(* IEC 61131-3 sources: guidance-for-physical-ai-production-designer-on-aws/source/plan2cell/examples/welding_cell_2_small/plc/codesys/robots/robot2/POU, 10 files *)

(* ---- FB_JointAngleEncoder.st ---- *)
(*
 * FB_JointAngleEncoder
 * Device simulator R2 (robot2), cell welding_cell_2_small. Generated by bt2plc 0.1.0.
 *
 * Encodes six KUKA robot joint angles (REAL degrees) into the VASS Option area
 * as scaled fixed-point INTs (0.02 deg per count, big-endian byte order).
 *
 * Encoding per encoding.md:
 *   count = ROUND(angle_deg / 0.02)   clamped to [-32768, +32767]
 *   Byte layout: big-endian (high byte first) in each 2-byte pair
 *
 * Output abyOption = Option area aVassInputData[16..27], 2 bytes per axis
 * (PLC_PRG copies it into the robot -> PLC telegram):
 *   abyOption[0-1]  = bytes 16-17 = A1,  abyOption[2-3]   = bytes 18-19 = A2,
 *   abyOption[4-5]  = bytes 20-21 = A3,  abyOption[6-7]   = bytes 22-23 = A4,
 *   abyOption[8-9]  = bytes 24-25 = A5,  abyOption[10-11] = bytes 26-27 = A6
 *)

FUNCTION_BLOCK FB_JointAngleEncoder
VAR_INPUT
    rA1_deg     : REAL := 0.0;      (* Axis 1 angle in degrees *)
    rA2_deg     : REAL := 0.0;      (* Axis 2 angle in degrees *)
    rA3_deg     : REAL := 0.0;      (* Axis 3 angle in degrees *)
    rA4_deg     : REAL := 0.0;      (* Axis 4 angle in degrees *)
    rA5_deg     : REAL := 0.0;      (* Axis 5 angle in degrees *)
    rA6_deg     : REAL := 0.0;      (* Axis 6 angle in degrees *)
END_VAR

VAR_OUTPUT
    (* Encoded INT values (for monitoring/debug) *)
    iA1_count   : INT;
    iA2_count   : INT;
    iA3_count   : INT;
    iA4_count   : INT;
    iA5_count   : INT;
    iA6_count   : INT;

    (* Option area bytes 16..27 of the robot -> PLC telegram, big-endian A1..A6 *)
    abyOption   : ARRAY[0..11] OF BYTE;
END_VAR

VAR CONSTANT
    SCALE_FACTOR    : REAL := 0.02;     (* degrees per count *)
    INV_SCALE       : REAL := 50.0;     (* 1/0.02 = 50, multiply for speed *)
    COUNT_MAX       : DINT := 32767;
    COUNT_MIN       : DINT := -32768;
END_VAR

VAR
    _arDeg      : ARRAY[1..6] OF REAL;
    _aiCount    : ARRAY[1..6] OF INT;
    _diTemp     : DINT;
    _wTemp      : WORD;
    _i          : INT;
END_VAR

(* ---- FB_PROFIsafe_Simulator.st ---- *)
(*
 * FB_PROFIsafe_Simulator
 * Device simulator R2 (robot2), cell welding_cell_2_small. Generated by bt2plc 0.1.0.
 *
 * Simulates the PROFIsafe protocol layer for the FDIO64 module (Slot 1).
 * In a real KUKA controller, the PROFIsafe stack handles CRC generation,
 * sequence counters, and watchdog monitoring.
 *
 * For simulation purposes, this FB:
 * - Monitors the safe output bytes from the PLC (abySafeOut = copy of GVL_IO.bySafeOut0..7)
 * - Provides a "communication OK" flag
 *
 * IMPORTANT: This does NOT provide real functional safety!
 * It only generates data patterns that allow the PLC's PROFIsafe stack
 * to accept the device as communicating. For real safety testing,
 * you need a certified PROFIsafe device or test equipment.
 *
 * PROFIsafe frame structure per IEC 61784-3-3:
 *   [User Data (8 bytes)] [Status/Control (1 byte)] [CRC (3 bytes)]
 *
 * Status byte bits (F_Input from device):
 *   Bit 0: Toggle bit (alternates each cycle)
 *   Bit 1: Reserved
 *   Bit 2: Data valid
 *   Bit 3-7: Reserved / Sequence counter
 *
 * Control byte bits (F_Output from controller):
 *   Bit 0: Toggle bit
 *   Bit 1: Activate device
 *   Bit 2: Reserved
 *   Bit 3-7: Reserved
 *)

FUNCTION_BLOCK FB_PROFIsafe_Simulator
VAR_INPUT
    bEnable         : BOOL := TRUE;
    dwF_Source_Add  : DWORD := DWORD#1;     (* F_Source_Add from parameterization *)
    dwF_Dest_Add    : DWORD := DWORD#1;     (* F_Dest_Add from parameterization *)
    tF_WD_Time      : TIME := T#500MS;      (* Watchdog time *)
    abySafeOut      : ARRAY[0..7] OF BYTE;  (* Safe outputs PLC -> robot (GVL_IO.bySafeOut0..7) *)
END_VAR

VAR_OUTPUT
    bCommOK         : BOOL;                 (* PROFIsafe communication established *)
    bDataValid      : BOOL;                 (* Safe data is valid *)
    bWatchdogError  : BOOL;                 (* Watchdog timeout *)
END_VAR

VAR
    _bToggleBit     : BOOL;                 (* Toggle bit for sequence *)
    _nSeqCounter    : BYTE;                 (* Sequence counter 0-31 *)
    _nCycleCount    : UDINT;                (* Absolute cycle counter *)

    (* Watchdog *)
    _tonWatchdog    : TON;
    _bPLCSafeActive : BOOL;

    (* CRC calculation helper *)
    _dwCrcSeed      : DWORD;
END_VAR

(* ---- FB_ProgramPlayer.st ---- *)
(*
 * FB_ProgramPlayer
 * Device simulator R2 (robot2), cell welding_cell_2_small, tree bt_1790934549_welding_cell_2_small. Generated by bt2plc 0.1.0.
 *
 * Plays the bt2plc robot program (GVL_Program) for PROD_FOLGE, or a blind joint
 * move to the home pose for HOME_FOLGE. Robot side of the zone protocol, per op k
 * with mask M = GVL_Program.aOps[k].dwZoneMask:
 *   1  wStep := k                          (also for M = 0)
 *   2  if M <> 0: REQUEST := M             (same call / telegram as wStep)
 *   3  if M <> 0: wait (GRANT AND M) = M
 *   4  start delay; trajectory (x rVelScale x override); hold
 *   5  if M <> 0: REQUEST := 0
 *   6  if M <> 0: wait (GRANT AND M) = 0   (4-phase, before the next REQUEST)
 *   7  next op; after the last op: bDone, wStep := 0 (same call)
 *
 * Timing: all times are REAL seconds accumulated from rDt (seconds per call, the
 * device task interval). Motion time advances by rDt * rRate * rVelScale, delay and
 * hold by rDt (the override does not scale dwell times). No TIME() / TON is used.
 * Zero-time transitions fall through within one call (at most N_MAX_TRANSITIONS),
 * but wStep changes at most once per call, so every step is visible to the head PLC.
 * Joints (deg) are linearly interpolated between waypoints and published as rA1..rA6_deg.
 * Abort (bAbort level while busy): REQUEST := 0, wStep := 0, the pose is held.
 * The robot powers up at GVL_Program.arHomeDeg.
 *)

FUNCTION_BLOCK FB_ProgramPlayer
VAR_INPUT
    bStart          : BOOL;                 (* Rising edge: start wJob *)
    wJob            : WORD;                 (* Folge to play: PROD_FOLGE or HOME_FOLGE *)
    bAbort          : BOOL;                 (* Level: stop / cancel / drives off / E-stop *)
    dwGrant         : DWORD;                (* Zone GRANT bits from the head PLC *)
    rRate           : REAL := 1.0;          (* Speed override factor (1.0 = 100 %) *)
    rDt             : REAL := 0.02;         (* Seconds per call (task interval) *)
END_VAR

VAR_OUTPUT
    eState          : E_PlayerState;        (* Current state *)
    bBusy           : BOOL;                 (* Program running *)
    bDone           : BOOL;                 (* Latched until next start *)
    bError          : BOOL;                 (* Latched until next start *)
    wErrorCode      : WORD;                 (* Error code, GVL_Program.ERR_xxx *)
    wWarningCode    : WORD;                 (* Warning code, GVL_Program.WARN_xxx, latched until next start *)
    wStep           : WORD;                 (* 1-based op index, 0 = none *)
    dwRequest       : DWORD;                (* Zone REQUEST bits to the head PLC *)
    bAtHome         : BOOL;                 (* All joints within R_AT_HOME_TOL_DEG of arHomeDeg *)
    rA1_deg         : REAL;                 (* Axis 1 angle *)
    rA2_deg         : REAL;                 (* Axis 2 angle *)
    rA3_deg         : REAL;                 (* Axis 3 angle *)
    rA4_deg         : REAL;                 (* Axis 4 angle *)
    rA5_deg         : REAL;                 (* Axis 5 angle *)
    rA6_deg         : REAL;                 (* Axis 6 angle *)
END_VAR

VAR CONSTANT
    N_MAX_TRANSITIONS : INT := 8;           (* Fall-through bound per call *)
END_VAR

VAR
    _eState         : E_PlayerState := E_PlayerState.PS_IDLE;
    _rtrigStart     : R_TRIG;
    _bFirstCall     : BOOL := TRUE;

    (* === Current op === *)
    _nOp            : INT;                  (* 1-based op index, 0 = HOME_FOLGE move *)
    _dwMask         : DWORD;                (* Zone mask of the current op *)
    _bHomeMove      : BOOL;                 (* Current move is a blind home move *)
    _nWp            : INT;                  (* Current waypoint segment start *)
    _nLast          : INT;                  (* Last waypoint of the current op, 0 = none *)
    _rVel           : REAL;                 (* Velocity scale of the current move *)

    (* === Time (s) === *)
    _rDtCall        : REAL;                 (* rDt limited to 0..1 s *)
    _rRateCall      : REAL;                 (* rRate limited to >= 0 *)
    _rT             : REAL;                 (* Motion time since move start *)
    _rTimer         : REAL;                 (* Delay / hold timer *)
    _rDur           : REAL;                 (* Duration of the blind home move *)
    _rAlpha         : REAL;                 (* Interpolation factor 0..1 *)
    _rSpan          : REAL;                 (* Waypoint segment duration *)

    (* === Pose (deg) === *)
    _arQ            : ARRAY[1..6] OF REAL;  (* Current joint angles *)
    _arQ0           : ARRAY[1..6] OF REAL;  (* Pose at the start of a blind home move *)
    _arQa           : ARRAY[1..6] OF REAL;  (* Segment start waypoint *)
    _arQb           : ARRAY[1..6] OF REAL;  (* Segment end waypoint *)

    (* === Fall-through === *)
    _nPass          : INT;
    _bAdvance       : BOOL;                 (* A transition happened in this pass *)
    _bStepSet       : BOOL;                 (* wStep changed in this call *)
    _bMoveDone      : BOOL;
    _i              : INT;
END_VAR

(* ---- FB_VASS_DeviceSimulator.st ---- *)
(*
 * FB_VASS_DeviceSimulator
 * Device simulator R2 (robot2, station kuka-robi2), cell welding_cell_2_small, tree bt_1790934549_welding_cell_2_small.
 * Generated by bt2plc 0.1.0.
 *
 * Simulates a KUKA KR C4 robot responding to VW VASS commands via PROFINET.
 *
 * This FB reads the PLC commands from its input images (PLC -> robot):
 *   aVassOutputData = copy of GVL_IO.aVassOutputData, abySafeOut = GVL_IO.bySafeOut0..7
 * and produces the robot status images (robot -> PLC):
 *   aVassInputData (bytes 16-27 = 0, the joint encoder fills them in PLC_PRG), abySafeIn.
 * PLC_PRG copies the images from / to GVL_IO; this FB never accesses GVL_IO.
 *
 * Job handshake (as the original simulator): drives on after 2 s, EXT mode, Ready,
 * JobRequest edge -> JobAck + job echo (clears ProgFinished), ProgStart edge -> start,
 * Stop/Cancel level -> stop, Reset held 500 ms -> clear error, gripper, speed override.
 * Job execution is delegated to FB_ProgramPlayer (GVL_Program):
 *   PROD_FOLGE: the bt2plc program; PLAN_ID (bytes PLAN_ID_BYTE..+1, latched at job accept)
 *               must equal GVL_Program.PLAN_ID at ProgStart, else ERR_PLAN_MISMATCH, no start.
 *   HOME_FOLGE: blind joint move to arHomeDeg (also on a HomeRequest [0].6 edge while Ready).
 *   other:      ERR_UNKNOWN_FOLGE, no start.
 * Zone protocol: wCurrentStep at bytes STEP_BYTE..+1, REQUEST DWORD LE at REQ_BYTE..+3,
 * GRANT DWORD LE read from bytes GRANT_BYTE..+3 (GVL_Program offsets).
 * At the end ProgRunning := FALSE, ProgFinished := TRUE and step := 0 in the same scan.
 *)

FUNCTION_BLOCK FB_VASS_DeviceSimulator
VAR_INPUT
    bEnable             : BOOL := TRUE;             (* Enable simulation *)
    wRobotID            : WORD := WORD#1;           (* Robot identification number 1-8 *)
    aVassOutputData     : ARRAY[0..31] OF BYTE;     (* VASS telegram PLC -> robot (GVL_IO.aVassOutputData) *)
    abySafeOut          : ARRAY[0..7] OF BYTE;      (* Safe outputs PLC -> robot (GVL_IO.bySafeOut0..7) *)
    rDt                 : REAL := 0.02;             (* Task interval in s (GVL_Program.R_TASK_S) *)
END_VAR

VAR_OUTPUT
    bActive             : BOOL;                     (* Simulator is active *)
    eCurrentMode        : E_RobotMode;              (* Current operating mode *)
    eProgramState       : E_ProgramState;           (* Current program state *)
    bSafetyOK           : BOOL;                     (* Safety system healthy *)
    aVassInputData      : ARRAY[0..31] OF BYTE;     (* VASS telegram robot -> PLC (bytes 16-27 = 0) *)
    abySafeIn           : ARRAY[0..7] OF BYTE;      (* Safe inputs robot -> PLC (GVL_IO.bySafeIn0..7) *)

    (* Joint angles from the program player (deg) *)
    rA1_deg             : REAL;
    rA2_deg             : REAL;
    rA3_deg             : REAL;
    rA4_deg             : REAL;
    rA5_deg             : REAL;
    rA6_deg             : REAL;

    (* Diagnostics *)
    wActiveJob          : WORD;                     (* Accepted job number (Folge) *)
    wCurrentStep        : WORD;                     (* Current op index, 0 = none *)
    wErrorCode          : WORD;                     (* Active error code *)
    dwRequest           : DWORD;                    (* Zone REQUEST bits sent to the head PLC *)
    dwGrant             : DWORD;                    (* Zone GRANT bits received from the head PLC *)
    ePlayerState        : E_PlayerState;            (* State of the program player *)
END_VAR

VAR
    (* === Internal Robot State === *)
    _bDrivesPowered     : BOOL;
    _bInExtMode         : BOOL;
    _bReady             : BOOL;
    _bError             : BOOL;
    _bProgRunning       : BOOL;
    _bAtHome            : BOOL := TRUE;
    _bInPosition        : BOOL := TRUE;
    _bProgFinished      : BOOL;
    _bJobAcknowledged   : BOOL;
    _bGripperClosed     : BOOL;
    _bPartPresent       : BOOL;
    _bPeriphReady       : BOOL := TRUE;

    _wActiveJob         : WORD;
    _wCurrentStep       : WORD;
    _wSpeed             : WORD := WORD#100;
    _wToolNr            : WORD := WORD#1;
    _wErrorCode         : WORD;
    _wWarningCode       : WORD;

    (* Simulated position (0.1mm units) *)
    _iPositionX         : INT := 5000;              (* 500.0 mm *)
    _iPositionY         : INT := 0;
    _iPositionZ         : INT := 10000;             (* 1000.0 mm *)

    (* === Safety State === *)
    _bSafe_DrivesOK     : BOOL := TRUE;
    _bSafe_Stopped      : BOOL := TRUE;
    _bSafe_EStopOK      : BOOL := TRUE;
    _bSafe_GatesClosed  : BOOL := TRUE;
    _bSafe_Fault        : BOOL;
    _bSafe_STO          : BOOL;
    _bSafe_SS1          : BOOL;

    (* PROFIsafe CRC simulation *)
    _bySafeTrailerStatus : BYTE;
    _nSafeCycleCount     : UDINT;

    (* === Timers === *)
    _tonDriveStartup    : TON;                      (* Simulate drive power-on delay *)
    _tonErrorReset      : TON;                      (* Simulate error reset delay *)
    _tonGripperAction   : TON;                      (* Simulate gripper open/close time *)

    (* === Edge Detection === *)
    _rtrigProgStart     : R_TRIG;
    _rtrigProgStop      : R_TRIG;
    _rtrigReset         : R_TRIG;
    _rtrigJobReq        : R_TRIG;
    _rtrigDrivesOn      : R_TRIG;
    _rtrigHome          : R_TRIG;
    _rtrigGripOpen      : R_TRIG;
    _rtrigGripClose     : R_TRIG;
    _rtrigSafeStop1     : R_TRIG;
    _rtrigSafeEStop     : R_TRIG;

    (* === Program player (bt2plc program / blind home) === *)
    _fbPlayer           : FB_ProgramPlayer;
    _bPlayerStart       : BOOL;                     (* Start pulse for the player *)
    _wPlayerJob         : WORD;                     (* Folge passed to the player *)
    _bStartOk           : BOOL;
    _wPlanId            : WORD;                     (* PLAN_ID latched at job accept *)
    _dwGrant            : DWORD;
    _dwRequest          : DWORD;
    _rRate              : REAL;                     (* Speed override factor *)
    _wPlayerWarning     : WORD;                     (* Last player warning (copy on change) *)

    (* === Decoded PLC commands (aVassOutputData bytes 0-1, abySafeOut byte 0) === *)
    _bCmdDrivesOn       : BOOL;                     (* [0].0 Drives on *)
    _bCmdProgStart      : BOOL;                     (* [0].1 Program start *)
    _bCmdProgStop       : BOOL;                     (* [0].2 Program stop *)
    _bCmdProgCancel     : BOOL;                     (* [0].3 Program cancel *)
    _bCmdModeExt        : BOOL;                     (* [0].4 EXT mode request *)
    _bCmdReset          : BOOL;                     (* [0].5 Reset *)
    _bCmdHome           : BOOL;                     (* [0].6 Home request *)
    _bCmdJobReq         : BOOL;                     (* [1].0 Job request *)
    _bCmdGripOpen       : BOOL;                     (* [1].1 Gripper open *)
    _bCmdGripClose      : BOOL;                     (* [1].2 Gripper close *)
    _bCmdSpeedOverride  : BOOL;                     (* [1].4 Apply speed override *)
    _bSafeCmdDriveEnable : BOOL;                    (* Safe [0].0 Drive enable *)
    _bSafeCmdEStop      : BOOL;                     (* Safe [0].1 External E-Stop *)
    _bSafeCmdSS1        : BOOL;                     (* Safe [0].2 Safe Stop 1 *)

    (* === Local working variables === *)
    _wRequestedJob      : WORD;
    _wSpeedCmd          : WORD;
    _nIdx               : INT;
    _i                  : INT;
END_VAR

(* ---- FB_JointAngleEncoder_Body.st ---- *)
(*
 * FB_JointAngleEncoder - Implementation
 *
 * Converts 6x REAL degree angles to scaled INT counts (0.02 deg per count)
 * and writes them big-endian into abyOption[0..11] (telegram bytes 16..27).
 *
 * Conversion:  count = ROUND(angle / 0.02)  clamped to INT range
 * Byte order:  Big-endian (high byte at lower address) per S7/PROFINET convention
 * Two's complement is formed in DINT (count + 65536 for negative counts), so no
 * bit operation is applied to a signed type.
 *)

_arDeg[1] := rA1_deg;
_arDeg[2] := rA2_deg;
_arDeg[3] := rA3_deg;
_arDeg[4] := rA4_deg;
_arDeg[5] := rA5_deg;
_arDeg[6] := rA6_deg;

FOR _i := 1 TO 6 DO
    (* === Scale and clamp === *)
    _diTemp := REAL_TO_DINT(LIMIT(REAL#-32768.0, _arDeg[_i] * INV_SCALE, REAL#32767.0));
    IF _diTemp > COUNT_MAX THEN _diTemp := COUNT_MAX; END_IF
    IF _diTemp < COUNT_MIN THEN _diTemp := COUNT_MIN; END_IF
    _aiCount[_i] := DINT_TO_INT(_diTemp);

    (* === Big-endian into the Option area: high byte first === *)
    IF _diTemp < 0 THEN
        _diTemp := _diTemp + 65536;
    END_IF
    _wTemp := DINT_TO_WORD(_diTemp);
    abyOption[2 * (_i - 1)] := WORD_TO_BYTE(SHR(_wTemp, 8));
    abyOption[2 * (_i - 1) + 1] := WORD_TO_BYTE(_wTemp AND WORD#16#FF);
END_FOR

iA1_count := _aiCount[1];
iA2_count := _aiCount[2];
iA3_count := _aiCount[3];
iA4_count := _aiCount[4];
iA5_count := _aiCount[5];
iA6_count := _aiCount[6];

(* ---- FB_PROFIsafe_Simulator_Body.st ---- *)
(*
 * FB_PROFIsafe_Simulator - Implementation
 * Works on the input image abySafeOut (PLC_PRG copies GVL_IO.bySafeOut0..7).
 *)

IF NOT bEnable THEN
    bCommOK := FALSE;
    bDataValid := FALSE;
    RETURN;
END_IF

IF _nCycleCount < UDINT#4000000000 THEN
    _nCycleCount := _nCycleCount + 1;
ELSE
    _nCycleCount := 0;
END_IF

(* ============================================================================
   MONITOR PLC SAFE OUTPUT DATA
   ============================================================================ *)
_bPLCSafeActive := (abySafeOut[0] <> BYTE#0) OR (abySafeOut[1] <> BYTE#0);

(* Watchdog *)
_tonWatchdog(IN := NOT _bPLCSafeActive, PT := tF_WD_Time);
bWatchdogError := _tonWatchdog.Q;

bCommOK := _bPLCSafeActive AND NOT bWatchdogError;
bDataValid := bCommOK;

(* ---- FB_ProgramPlayer_Body.st ---- *)
(*
 * FB_ProgramPlayer - Implementation
 *)

(* ============================================================================
   INIT - the robot powers up at the home pose
   ============================================================================ *)
IF _bFirstCall THEN
    FOR _i := 1 TO 6 DO
        _arQ[_i] := GVL_Program.arHomeDeg[_i];
    END_FOR
    _bFirstCall := FALSE;
END_IF

_rDtCall := LIMIT(0.0, rDt, 1.0);
_rRateCall := MAX(rRate, 0.0);
_rtrigStart(CLK := bStart);

(* ============================================================================
   ABORT - stop / cancel / drives off / E-stop: REQUEST := 0, wStep := 0, hold pose
   ============================================================================ *)
IF bAbort AND bBusy THEN
    _eState := E_PlayerState.PS_IDLE;
    bBusy := FALSE;
    wStep := WORD#0;
    dwRequest := DWORD#0;
END_IF

(* ============================================================================
   CLOCK - advance the timer of the state that is active at the start of the call
   (a state entered during this call starts counting with the next call)
   ============================================================================ *)
IF _eState = E_PlayerState.PS_DELAY OR _eState = E_PlayerState.PS_HOLD THEN
    _rTimer := _rTimer + _rDtCall;
ELSIF _eState = E_PlayerState.PS_MOVE THEN
    _rT := _rT + _rDtCall * _rRateCall * _rVel;
END_IF

(* ============================================================================
   START
   ============================================================================ *)
IF _rtrigStart.Q AND NOT bBusy AND NOT bAbort THEN
    bDone := FALSE;
    bError := FALSE;
    wErrorCode := WORD#0;
    wWarningCode := WORD#0;
    wStep := WORD#0;
    dwRequest := DWORD#0;
    _nOp := 0;
    _dwMask := DWORD#0;
    _rT := 0.0;
    _rTimer := 0.0;
    IF wJob = GVL_Program.HOME_FOLGE THEN
        (* Blind joint move from the current pose to arHomeDeg: no step, no zones *)
        FOR _i := 1 TO 6 DO
            _arQ0[_i] := _arQ[_i];
        END_FOR
        _bHomeMove := TRUE;
        _nLast := 0;
        _rVel := 1.0;
        _rDur := GVL_Program.R_HOME_S;
        bBusy := TRUE;
        _eState := E_PlayerState.PS_MOVE;
    ELSIF wJob = GVL_Program.PROD_FOLGE AND GVL_Program.N_OPS > 0 THEN
        bBusy := TRUE;
        _eState := E_PlayerState.PS_NEXT_OP;
    ELSE
        wErrorCode := GVL_Program.ERR_UNKNOWN_FOLGE;
        _eState := E_PlayerState.PS_ERROR;
    END_IF
END_IF

(* ============================================================================
   STATE MACHINE - falls through zero-time transitions (bounded)
   ============================================================================ *)
_bStepSet := FALSE;
FOR _nPass := 1 TO N_MAX_TRANSITIONS DO
    _bAdvance := FALSE;

    CASE _eState OF

    E_PlayerState.PS_IDLE:
        bBusy := FALSE;
        wStep := WORD#0;
        dwRequest := DWORD#0;

    E_PlayerState.PS_NEXT_OP:
        (* wStep changes at most once per call: the head checks step + 1 per telegram *)
        IF NOT _bStepSet THEN
            _nOp := _nOp + 1;
            IF _nOp > GVL_Program.N_OPS THEN
                _eState := E_PlayerState.PS_DONE;
            ELSE
                wStep := INT_TO_WORD(_nOp);
                _bStepSet := TRUE;
                _dwMask := GVL_Program.aOps[_nOp].dwZoneMask;
                IF _dwMask <> DWORD#0 THEN
                    dwRequest := _dwMask;           (* same telegram as wStep *)
                    _eState := E_PlayerState.PS_WAIT_GRANT;
                ELSE
                    _rTimer := 0.0;
                    _eState := E_PlayerState.PS_DELAY;
                END_IF
            END_IF
            _bAdvance := TRUE;
        END_IF

    E_PlayerState.PS_WAIT_GRANT:
        IF (dwGrant AND _dwMask) = _dwMask THEN
            _rTimer := 0.0;
            _eState := E_PlayerState.PS_DELAY;
            _bAdvance := TRUE;
        END_IF

    E_PlayerState.PS_DELAY:
        IF _rTimer >= GVL_Program.aOps[_nOp].rDelay_s THEN
            (* Begin the motion of op _nOp *)
            _rT := 0.0;
            _rVel := GVL_Program.aOps[_nOp].rVelScale;
            IF _rVel <= 0.0 THEN
                _rVel := 1.0;
            END_IF
            _bHomeMove := GVL_Program.aOps[_nOp].bBlindHome;
            IF _bHomeMove THEN
                FOR _i := 1 TO 6 DO
                    _arQ0[_i] := _arQ[_i];
                END_FOR
                _rDur := GVL_Program.R_HOME_S;
                _nLast := 0;
            ELSE
                _nWp := GVL_Program.aOps[_nOp].nFirstWp;
                _nLast := GVL_Program.aOps[_nOp].nLastWp;
                IF _nWp < 1 OR _nLast < _nWp OR _nLast > GVL_Program.N_WP THEN
                    _nLast := 0;                    (* no valid trajectory: zero-length move *)
                ELSE
                    (* Start deviation: the trajectory should start at the current pose *)
                    _arQa[1] := GVL_Program.aWp[_nWp].rA1;
                    _arQa[2] := GVL_Program.aWp[_nWp].rA2;
                    _arQa[3] := GVL_Program.aWp[_nWp].rA3;
                    _arQa[4] := GVL_Program.aWp[_nWp].rA4;
                    _arQa[5] := GVL_Program.aWp[_nWp].rA5;
                    _arQa[6] := GVL_Program.aWp[_nWp].rA6;
                    FOR _i := 1 TO 6 DO
                        IF ABS(_arQ[_i] - _arQa[_i]) > GVL_Program.R_START_TOL_DEG THEN
                            wWarningCode := GVL_Program.WARN_START_DEVIATION;
                        END_IF
                    END_FOR
                END_IF
            END_IF
            _eState := E_PlayerState.PS_MOVE;
            _bAdvance := TRUE;
        END_IF

    E_PlayerState.PS_MOVE:
        _bMoveDone := FALSE;
        IF _bHomeMove THEN
            (* Blind joint move: linear in joint space over R_HOME_S *)
            IF _rDur > 0.0 THEN
                _rAlpha := LIMIT(0.0, _rT / _rDur, 1.0);
            ELSE
                _rAlpha := 1.0;
            END_IF
            FOR _i := 1 TO 6 DO
                _arQ[_i] := _arQ0[_i] + _rAlpha * (GVL_Program.arHomeDeg[_i] - _arQ0[_i]);
            END_FOR
            _bMoveDone := _rAlpha >= 1.0;
        ELSIF _nLast < 1 THEN
            _bMoveDone := TRUE;
        ELSE
            (* Trajectory: find the segment [_nWp, _nWp + 1] that contains _rT *)
            WHILE _nWp < _nLast DO
                IF GVL_Program.aWp[_nWp + 1].rT <= _rT THEN
                    _nWp := _nWp + 1;
                ELSE
                    EXIT;
                END_IF
            END_WHILE
            _arQa[1] := GVL_Program.aWp[_nWp].rA1;
            _arQa[2] := GVL_Program.aWp[_nWp].rA2;
            _arQa[3] := GVL_Program.aWp[_nWp].rA3;
            _arQa[4] := GVL_Program.aWp[_nWp].rA4;
            _arQa[5] := GVL_Program.aWp[_nWp].rA5;
            _arQa[6] := GVL_Program.aWp[_nWp].rA6;
            IF _nWp >= _nLast THEN
                FOR _i := 1 TO 6 DO
                    _arQ[_i] := _arQa[_i];
                END_FOR
                _bMoveDone := TRUE;
            ELSE
                _arQb[1] := GVL_Program.aWp[_nWp + 1].rA1;
                _arQb[2] := GVL_Program.aWp[_nWp + 1].rA2;
                _arQb[3] := GVL_Program.aWp[_nWp + 1].rA3;
                _arQb[4] := GVL_Program.aWp[_nWp + 1].rA4;
                _arQb[5] := GVL_Program.aWp[_nWp + 1].rA5;
                _arQb[6] := GVL_Program.aWp[_nWp + 1].rA6;
                _rSpan := GVL_Program.aWp[_nWp + 1].rT - GVL_Program.aWp[_nWp].rT;
                IF _rSpan > 0.0 THEN
                    _rAlpha := LIMIT(0.0, (_rT - GVL_Program.aWp[_nWp].rT) / _rSpan, 1.0);
                ELSE
                    _rAlpha := 1.0;
                END_IF
                FOR _i := 1 TO 6 DO
                    _arQ[_i] := _arQa[_i] + _rAlpha * (_arQb[_i] - _arQa[_i]);
                END_FOR
            END_IF
        END_IF
        IF _bMoveDone THEN
            IF _nOp = 0 THEN
                _eState := E_PlayerState.PS_DONE;   (* HOME_FOLGE finished *)
            ELSE
                _rTimer := 0.0;
                _eState := E_PlayerState.PS_HOLD;
            END_IF
            _bAdvance := TRUE;
        END_IF

    E_PlayerState.PS_HOLD:
        IF _rTimer >= GVL_Program.aOps[_nOp].rHold_s THEN
            IF _dwMask <> DWORD#0 THEN
                dwRequest := DWORD#0;
                _eState := E_PlayerState.PS_WAIT_RELEASE;
            ELSE
                _eState := E_PlayerState.PS_NEXT_OP;
            END_IF
            _bAdvance := TRUE;
        END_IF

    E_PlayerState.PS_WAIT_RELEASE:
        (* 4-phase: the GRANT must drop before the next REQUEST *)
        IF (dwGrant AND _dwMask) = DWORD#0 THEN
            _eState := E_PlayerState.PS_NEXT_OP;
            _bAdvance := TRUE;
        END_IF

    E_PlayerState.PS_DONE:
        bBusy := FALSE;
        bDone := TRUE;
        wStep := WORD#0;
        dwRequest := DWORD#0;
        _eState := E_PlayerState.PS_IDLE;

    E_PlayerState.PS_ERROR:
        bBusy := FALSE;
        bError := TRUE;
        wStep := WORD#0;
        dwRequest := DWORD#0;
        _eState := E_PlayerState.PS_IDLE;

    END_CASE

    IF NOT _bAdvance THEN
        EXIT;
    END_IF
END_FOR

(* ============================================================================
   PUBLISH
   ============================================================================ *)
bAtHome := TRUE;
FOR _i := 1 TO 6 DO
    IF ABS(_arQ[_i] - GVL_Program.arHomeDeg[_i]) > GVL_Program.R_AT_HOME_TOL_DEG THEN
        bAtHome := FALSE;
    END_IF
END_FOR
rA1_deg := _arQ[1];
rA2_deg := _arQ[2];
rA3_deg := _arQ[3];
rA4_deg := _arQ[4];
rA5_deg := _arQ[5];
rA6_deg := _arQ[6];
eState := _eState;

(* ---- FB_VASS_DeviceSimulator_Body.st ---- *)
(*
 * FB_VASS_DeviceSimulator - Implementation
 *
 * Reads commands from aVassOutputData (PLC -> Robot, 32 bytes) and abySafeOut (8 bytes).
 * Writes status to aVassInputData (Robot -> PLC, 32 bytes) and abySafeIn (8 bytes).
 *)

IF NOT bEnable THEN
    bActive := FALSE;
    RETURN;
END_IF

bActive := TRUE;

(* ============================================================================
   SECTION 1: READ PLC COMMANDS from aVassOutputData[0..31]
   Byte 0-1 = Control word, Byte 2-3 = Job number, PLAN_ID / GRANT per GVL_Program
   ============================================================================ *)

(* Decode the control bits into BOOLs (a bare bit access is never passed as a call argument) *)
_bCmdDrivesOn       := aVassOutputData[0].0;
_bCmdProgStart      := aVassOutputData[0].1;
_bCmdProgStop       := aVassOutputData[0].2;
_bCmdProgCancel     := aVassOutputData[0].3;
_bCmdModeExt        := aVassOutputData[0].4;
_bCmdReset          := aVassOutputData[0].5;
_bCmdHome           := aVassOutputData[0].6;
_bCmdJobReq         := aVassOutputData[1].0;
_bCmdGripOpen       := aVassOutputData[1].1;
_bCmdGripClose      := aVassOutputData[1].2;
_bCmdSpeedOverride  := aVassOutputData[1].4;
_bSafeCmdDriveEnable := abySafeOut[0].0;
_bSafeCmdEStop      := abySafeOut[0].1;
_bSafeCmdSS1        := abySafeOut[0].2;

(* Edge detection on control signals - output byte 0 *)
_rtrigDrivesOn(CLK  := _bCmdDrivesOn);
_rtrigProgStart(CLK := _bCmdProgStart);
_rtrigProgStop(CLK  := _bCmdProgStop);
_rtrigReset(CLK     := _bCmdReset);
_rtrigHome(CLK      := _bCmdHome);

(* Output byte 1 *)
_rtrigJobReq(CLK    := _bCmdJobReq);
_rtrigGripOpen(CLK  := _bCmdGripOpen);
_rtrigGripClose(CLK := _bCmdGripClose);

(* Safety edge detection from safe output byte 0 *)
_rtrigSafeStop1(CLK := _bSafeCmdSS1);
_rtrigSafeEStop(CLK := _bSafeCmdEStop);

(* Requested job number: bytes 2-3 WORD LE, or byte 2 only (GVL_Program.JOB_NUMBER_BYTE) *)
IF GVL_Program.JOB_NUMBER_BYTE THEN
    _wRequestedJob := BYTE_TO_WORD(aVassOutputData[2]);
ELSE
    _wRequestedJob := BYTE_TO_WORD(aVassOutputData[2])
                      OR SHL(BYTE_TO_WORD(aVassOutputData[3]), 8);
END_IF

(* Zone GRANT: DWORD LE at bytes GVL_Program.GRANT_BYTE..+3 *)
_nIdx := GVL_Program.GRANT_BYTE;
_dwGrant := BYTE_TO_DWORD(aVassOutputData[_nIdx])
            OR SHL(BYTE_TO_DWORD(aVassOutputData[_nIdx + 1]), 8)
            OR SHL(BYTE_TO_DWORD(aVassOutputData[_nIdx + 2]), 16)
            OR SHL(BYTE_TO_DWORD(aVassOutputData[_nIdx + 3]), 24);

(* ============================================================================
   SECTION 2: SAFETY LOGIC (PROFIsafe Slot 1)
   Reads abySafeOut, status is written to abySafeIn in section 4
   ============================================================================ *)

(* Process safe outputs from PLC - byte 0 *)
_bSafe_DrivesOK := _bSafeCmdDriveEnable AND _bSafe_EStopOK AND NOT _bSafe_Fault;

(* E-Stop handling *)
IF _bSafeCmdEStop THEN  (* External E-Stop *)
    _bSafe_EStopOK := FALSE;
    _bSafe_STO := TRUE;
    _bDrivesPowered := FALSE;
    _bProgRunning := FALSE;
    eProgramState := E_ProgramState.PRG_STOPPED;
END_IF

(* Safe Stop 1 request *)
IF _bSafeCmdSS1 AND _bProgRunning THEN
    _bSafe_SS1 := TRUE;
    _bProgRunning := FALSE;
    _bSafe_Stopped := TRUE;
    eProgramState := E_ProgramState.PRG_STOPPED;
END_IF

(* Recovery from safety state *)
IF NOT _bSafeCmdEStop AND NOT _bSafeCmdSS1 THEN
    IF _bCmdReset THEN  (* Reset bit *)
        _bSafe_EStopOK := TRUE;
        _bSafe_STO := FALSE;
        _bSafe_SS1 := FALSE;
        _bSafe_Stopped := FALSE;
        _bSafe_Fault := FALSE;
    END_IF
END_IF

(* Overall safety status *)
bSafetyOK := _bSafe_DrivesOK AND _bSafe_EStopOK AND _bSafe_GatesClosed AND NOT _bSafe_Fault;
_bSafe_GatesClosed := TRUE; (* Always closed in simulation *)

(* ============================================================================
   SECTION 3: STANDARD I/O LOGIC (VASS Telegram Slot 2)
   ============================================================================ *)

(* --- Drive Power Control --- *)
_tonDriveStartup(IN := _bCmdDrivesOn AND bSafetyOK AND NOT _bDrivesPowered, PT := T#2S);
IF _tonDriveStartup.Q THEN
    _bDrivesPowered := TRUE;
    _bSafe_Stopped := FALSE;
END_IF

IF NOT _bCmdDrivesOn OR NOT bSafetyOK THEN
    _bDrivesPowered := FALSE;
    _bProgRunning := FALSE;
    IF eProgramState = E_ProgramState.PRG_RUNNING THEN
        eProgramState := E_ProgramState.PRG_STOPPED;
    END_IF
END_IF

(* --- Mode Control --- *)
_bInExtMode := _bCmdModeExt AND _bDrivesPowered AND bSafetyOK;
IF _bInExtMode THEN
    eCurrentMode := E_RobotMode.MODE_EXT;
ELSE
    eCurrentMode := E_RobotMode.MODE_T1;
END_IF

(* --- Ready State --- *)
_bReady := _bDrivesPowered
           AND _bInExtMode
           AND NOT _bError
           AND NOT _bProgRunning
           AND bSafetyOK;

(* --- Warning reset: any Reset edge clears a pending warning (no error needed) --- *)
IF _rtrigReset.Q THEN
    _wWarningCode := WORD#0;
END_IF

(* --- Error Reset (Reset held 500 ms) --- *)
_tonErrorReset(IN := _bCmdReset AND _bError, PT := T#500MS);
IF _tonErrorReset.Q THEN
    _bError := FALSE;
    _wErrorCode := WORD#0;
    _wWarningCode := WORD#0;
    IF eProgramState = E_ProgramState.PRG_ERROR THEN
        eProgramState := E_ProgramState.PRG_IDLE;
    END_IF
END_IF

(* --- Job Request Handling --- *)
IF _rtrigJobReq.Q AND _bReady THEN
    _wActiveJob := _wRequestedJob;
    _bJobAcknowledged := TRUE;
    _bProgFinished := FALSE;
    (* PLAN_ID: WORD LE at bytes GVL_Program.PLAN_ID_BYTE..+1 (production job only) *)
    _nIdx := GVL_Program.PLAN_ID_BYTE;
    _wPlanId := BYTE_TO_WORD(aVassOutputData[_nIdx])
                OR SHL(BYTE_TO_WORD(aVassOutputData[_nIdx + 1]), 8);
END_IF

IF NOT _bCmdJobReq THEN
    _bJobAcknowledged := FALSE;
END_IF

(* --- Program Start --- *)
_bStartOk := FALSE;
IF _rtrigProgStart.Q AND _bReady AND _wActiveJob <> WORD#0 THEN
    _wPlayerJob := _wActiveJob;
    IF _wActiveJob = GVL_Program.HOME_FOLGE THEN
        _bStartOk := TRUE;
    ELSIF _wActiveJob = GVL_Program.PROD_FOLGE AND GVL_Program.N_OPS > 0 THEN
        IF _wPlanId = GVL_Program.PLAN_ID THEN
            _bStartOk := TRUE;
        ELSE
            _bError := TRUE;
            _wErrorCode := GVL_Program.ERR_PLAN_MISMATCH;
            eProgramState := E_ProgramState.PRG_ERROR;
        END_IF
    ELSE
        _bError := TRUE;
        _wErrorCode := GVL_Program.ERR_UNKNOWN_FOLGE;
        eProgramState := E_ProgramState.PRG_ERROR;
    END_IF
ELSIF _rtrigHome.Q AND _bReady AND NOT _bAtHome THEN
    (* HomeRequest [0].6 edge while Ready: behaves like HOME_FOLGE *)
    _wPlayerJob := GVL_Program.HOME_FOLGE;
    _bStartOk := TRUE;
END_IF

IF _bStartOk THEN
    _bProgRunning := TRUE;
    _bProgFinished := FALSE;
    _bInPosition := FALSE;
    _bSafe_Stopped := FALSE;
    _bPlayerStart := TRUE;
    eProgramState := E_ProgramState.PRG_RUNNING;
END_IF

(* --- Program Stop/Cancel (level) --- *)
IF (_bCmdProgStop OR _bCmdProgCancel) AND _bProgRunning THEN
    _bProgRunning := FALSE;
    _bProgFinished := FALSE;
    _bInPosition := TRUE;
    eProgramState := E_ProgramState.PRG_STOPPED;
END_IF

(* --- Program Execution: FB_ProgramPlayer --- *)
(* Any stop path above (Stop/Cancel, drives off, E-stop, SS1) aborts the player in this scan:
   REQUEST := 0, step := 0, the pose is held. *)
_rRate := UINT_TO_REAL(WORD_TO_UINT(_wSpeed)) / 100.0;
_fbPlayer(
    bStart  := _bPlayerStart,
    wJob    := _wPlayerJob,
    bAbort  := NOT _bProgRunning,
    dwGrant := _dwGrant,
    rRate   := _rRate,
    rDt     := rDt
);
_bPlayerStart := FALSE;

IF _bProgRunning THEN
    IF _fbPlayer.bError THEN
        _bProgRunning := FALSE;
        _bError := TRUE;
        _wErrorCode := _fbPlayer.wErrorCode;
        eProgramState := E_ProgramState.PRG_ERROR;
    ELSIF _fbPlayer.bDone THEN
        (* Same scan as step := 0: ProgRunning drops and ProgFinished rises together *)
        _bProgRunning := FALSE;
        _bProgFinished := TRUE;
        _bInPosition := TRUE;
        eProgramState := E_ProgramState.PRG_FINISHED;
    END_IF
END_IF

_wCurrentStep := _fbPlayer.wStep;
_dwRequest := _fbPlayer.dwRequest;
_bAtHome := _fbPlayer.bAtHome;

(* Player warnings are copied on change, so an error reset clears them *)
IF _fbPlayer.wWarningCode <> _wPlayerWarning THEN
    _wPlayerWarning := _fbPlayer.wWarningCode;
    IF _wPlayerWarning <> WORD#0 THEN
        _wWarningCode := _wPlayerWarning;
    END_IF
END_IF

(* --- Gripper Simulation --- *)
_tonGripperAction(IN := _bCmdGripClose AND NOT _bGripperClosed, PT := T#500MS);
IF _tonGripperAction.Q THEN
    _bGripperClosed := TRUE;
    _bPartPresent := TRUE;
END_IF

IF _bCmdGripOpen THEN
    _bGripperClosed := FALSE;
    _bPartPresent := FALSE;
END_IF

(* --- Speed Override (bytes 8-9 WORD LE, applied with [1].4) --- *)
_wSpeedCmd := BYTE_TO_WORD(aVassOutputData[8]) OR SHL(BYTE_TO_WORD(aVassOutputData[9]), 8);
IF _bCmdSpeedOverride AND WORD_TO_UINT(_wSpeedCmd) > 0 AND WORD_TO_UINT(_wSpeedCmd) <= 100 THEN
    _wSpeed := _wSpeedCmd;
END_IF

(* ============================================================================
   SECTION 4: WRITE SAFETY STATUS to abySafeIn[0..7]
   ============================================================================ *)

(* Byte 0: Safe drive/motion status *)
abySafeIn[0].0 := _bSafe_DrivesOK;
abySafeIn[0].1 := _bSafe_Stopped;
abySafeIn[0].2 := FALSE; (* Reduced speed *)
abySafeIn[0].3 := NOT _bSafe_Fault; (* Axis monitor OK *)
abySafeIn[0].4 := TRUE;  (* Tool monitor OK *)
abySafeIn[0].5 := TRUE;  (* Workspace OK *)
abySafeIn[0].6 := FALSE;
abySafeIn[0].7 := FALSE;

(* Byte 1: Gate/protection status *)
abySafeIn[1].0 := _bSafe_GatesClosed;  (* Gate 1 *)
abySafeIn[1].1 := _bSafe_GatesClosed;  (* Gate 2 *)
abySafeIn[1].2 := _bSafe_GatesClosed;  (* Gate 3 *)
abySafeIn[1].3 := TRUE;   (* Light curtain OK *)
abySafeIn[1].4 := _bSafe_EStopOK;
abySafeIn[1].5 := FALSE;  (* Enabling device *)
abySafeIn[1].6 := TRUE;   (* Operator safe *)
abySafeIn[1].7 := FALSE;

(* Byte 2: Extended safe functions *)
abySafeIn[2].0 := _bSafe_STO;
abySafeIn[2].1 := _bSafe_SS1;
abySafeIn[2].2 := FALSE;  (* SS2 *)
abySafeIn[2].3 := _bSafe_Stopped AND NOT _bSafe_STO;  (* SOS *)
abySafeIn[2].4 := FALSE;  (* SLS *)
abySafeIn[2].5 := FALSE;  (* SLP *)
abySafeIn[2].6 := FALSE;
abySafeIn[2].7 := _bSafe_Fault;

(* Bytes 3-7: zero *)
abySafeIn[3] := BYTE#0;
abySafeIn[4] := BYTE#0;
abySafeIn[5] := BYTE#0;
abySafeIn[6] := BYTE#0;
abySafeIn[7] := BYTE#0;

(* ============================================================================
   SECTION 5: WRITE VASS STATUS to aVassInputData[0..31]
   ============================================================================ *)

(* Unused bytes are zero; bytes 16-27 (joint angles) are filled by PLC_PRG *)
FOR _i := 0 TO 31 DO
    aVassInputData[_i] := BYTE#0;
END_FOR

(* Status Word - Byte 0 *)
aVassInputData[0].0 := _bDrivesPowered;
aVassInputData[0].1 := _bProgRunning;
aVassInputData[0].2 := _bAtHome;
aVassInputData[0].3 := _bInPosition;
aVassInputData[0].4 := _bInExtMode;
aVassInputData[0].5 := _bReady;
aVassInputData[0].6 := _bError;
aVassInputData[0].7 := _wWarningCode <> WORD#0;

(* Status Word - Byte 1 *)
aVassInputData[1].0 := _bSafe_GatesClosed;
aVassInputData[1].1 := _bSafe_EStopOK;
aVassInputData[1].2 := _bProgFinished;
aVassInputData[1].3 := _bJobAcknowledged;
aVassInputData[1].4 := _bGripperClosed;
aVassInputData[1].5 := _bPartPresent;
aVassInputData[1].6 := TRUE;  (* Periph ready *)
aVassInputData[1].7 := FALSE; (* Maint not required *)

(* Active job number echo - Bytes 2-3 (byte 2 only in byte mode, byte 3 = 0) *)
aVassInputData[2] := WORD_TO_BYTE(_wActiveJob AND WORD#16#FF);
IF NOT GVL_Program.JOB_NUMBER_BYTE THEN
    aVassInputData[3] := WORD_TO_BYTE(SHR(_wActiveJob, 8));
END_IF

(* Speed actual - Bytes 6-7 *)
aVassInputData[6] := WORD_TO_BYTE(_wSpeed AND WORD#16#FF);
aVassInputData[7] := WORD_TO_BYTE(SHR(_wSpeed, 8));

(* Tool number - Bytes 8-9 *)
aVassInputData[8] := WORD_TO_BYTE(_wToolNr AND WORD#16#FF);
aVassInputData[9] := WORD_TO_BYTE(SHR(_wToolNr, 8));

(* Error code - Bytes 10-11 *)
aVassInputData[10] := WORD_TO_BYTE(_wErrorCode AND WORD#16#FF);
aVassInputData[11] := WORD_TO_BYTE(SHR(_wErrorCode, 8));

(* Warning code - Bytes 12-13 *)
aVassInputData[12] := WORD_TO_BYTE(_wWarningCode AND WORD#16#FF);
aVassInputData[13] := WORD_TO_BYTE(SHR(_wWarningCode, 8));

(* Position X - Bytes 14-15 *)
aVassInputData[14] := WORD_TO_BYTE(INT_TO_WORD(_iPositionX) AND WORD#16#FF);
aVassInputData[15] := WORD_TO_BYTE(SHR(INT_TO_WORD(_iPositionX), 8));

(* Bytes 16-27: A129_224_Option area - RESERVED for the joint angle encoder
   (PLC_PRG -> fbJointEncoder, 6x INT big-endian = A1..A6 at 0.02 deg/count) *)

(* Current step (op index) - WORD LE at bytes GVL_Program.STEP_BYTE..+1 *)
_nIdx := GVL_Program.STEP_BYTE;
aVassInputData[_nIdx] := WORD_TO_BYTE(_wCurrentStep AND WORD#16#FF);
aVassInputData[_nIdx + 1] := WORD_TO_BYTE(SHR(_wCurrentStep, 8));

(* Zone REQUEST - DWORD LE at bytes GVL_Program.REQ_BYTE..+3 *)
_nIdx := GVL_Program.REQ_BYTE;
aVassInputData[_nIdx] := DWORD_TO_BYTE(_dwRequest AND DWORD#16#FF);
aVassInputData[_nIdx + 1] := DWORD_TO_BYTE(SHR(_dwRequest, 8) AND DWORD#16#FF);
aVassInputData[_nIdx + 2] := DWORD_TO_BYTE(SHR(_dwRequest, 16) AND DWORD#16#FF);
aVassInputData[_nIdx + 3] := DWORD_TO_BYTE(SHR(_dwRequest, 24));

(* ============================================================================
   SECTION 6: OUTPUTS (joint angles, diagnostics)
   ============================================================================ *)
rA1_deg := _fbPlayer.rA1_deg;
rA2_deg := _fbPlayer.rA2_deg;
rA3_deg := _fbPlayer.rA3_deg;
rA4_deg := _fbPlayer.rA4_deg;
rA5_deg := _fbPlayer.rA5_deg;
rA6_deg := _fbPlayer.rA6_deg;

wActiveJob := _wActiveJob;
wCurrentStep := _wCurrentStep;
wErrorCode := _wErrorCode;
dwRequest := _dwRequest;
dwGrant := _dwGrant;
ePlayerState := _fbPlayer.eState;

(* ---- PLC_PRG.st ---- *)
(*
 * PLC_PRG
 * Main program of the KUKA VASS device simulator R2 (robot2, station kuka-robi2),
 * cell welding_cell_2_small, tree bt_1790934549_welding_cell_2_small. Generated by bt2plc 0.1.0.
 *
 * I/O Flow (only this program accesses GVL_IO; FBs work on the local images):
 *   PLC -> PROFINET -> GVL_IO.aVassOutputData[0..31] -> aVassOutputData -> simulator reads commands
 *   PLC -> PROFIsafe -> GVL_IO.bySafeOut0..7         -> abySafeOut      -> simulator reads safe cmds
 *   simulator -> aVassInputData -> GVL_IO.aVassInputData[0..31] (whole array) -> PROFINET -> PLC
 *   simulator -> abySafeIn      -> GVL_IO.bySafeIn0..7 (scalars)              -> PROFIsafe -> PLC
 *
 * Joint angle flow:
 *   FB_ProgramPlayer (inside fbVassSimulator, GVL_Program) -> FB_JointAngleEncoder
 *   -> aVassInputData[16..27]
 *
 * Task: MainTask, interval GVL_Program.R_TASK_S (passed to the player as rDt)
 *)

PROGRAM PLC_PRG
VAR
    (* Main simulator instances *)
    fbVassSimulator         : FB_VASS_DeviceSimulator;
    fbSafetySimulator       : FB_PROFIsafe_Simulator;

    (* Joint angle encoding *)
    fbJointEncoder          : FB_JointAngleEncoder;

    (* === Configuration === *)
    bSimulatorEnable        : BOOL := TRUE;     (* Enable/disable simulator *)

    (* PROFIsafe parameters *)
    dwF_Source_Add          : DWORD := DWORD#1;
    dwF_Dest_Add            : DWORD := DWORD#1;
    tF_WD_Time              : TIME := T#500MS;

    (* === Local I/O images (copied from / to GVL_IO as a whole) === *)
    aVassOutputData         : ARRAY[0..31] OF BYTE;     (* PLC -> robot *)
    aVassInputData          : ARRAY[0..31] OF BYTE;     (* robot -> PLC *)
    abySafeOut              : ARRAY[0..7] OF BYTE;      (* PLC -> robot, GVL_IO.bySafeOut0..7 *)
    abySafeIn               : ARRAY[0..7] OF BYTE;      (* robot -> PLC, GVL_IO.bySafeIn0..7 *)

    (* === Diagnostic outputs === *)
    bSimActive              : BOOL;
    eMode                   : E_RobotMode;
    eProgState              : E_ProgramState;
    bSafetyHealthy          : BOOL;
    bSafeCommOK             : BOOL;
    wActiveJob              : WORD;
    wCurrentStep            : WORD;
    dwRequest               : DWORD;
    dwGrant                 : DWORD;
    ePlayerState            : E_PlayerState;

    (* Joint angle monitor (decoded back for verification) *)
    rMonitor_A1_deg         : REAL;
    rMonitor_A2_deg         : REAL;
    rMonitor_A3_deg         : REAL;
    rMonitor_A4_deg         : REAL;
    rMonitor_A5_deg         : REAL;
    rMonitor_A6_deg         : REAL;

    (* === Test/Debug signals === *)
    bTest_InjectError       : BOOL;
    bTest_InjectSafetyFault : BOOL;
    wTest_ErrorCode         : WORD := WORD#16#0010;

    _i                      : INT;
END_VAR

(* ---- PLC_PRG_Body.st ---- *)
(* ============================================================================
   INPUTS: copy the head PLC commands into the local images
   ============================================================================ *)
aVassOutputData := GVL_IO.aVassOutputData;
abySafeOut[0] := GVL_IO.bySafeOut0;
abySafeOut[1] := GVL_IO.bySafeOut1;
abySafeOut[2] := GVL_IO.bySafeOut2;
abySafeOut[3] := GVL_IO.bySafeOut3;
abySafeOut[4] := GVL_IO.bySafeOut4;
abySafeOut[5] := GVL_IO.bySafeOut5;
abySafeOut[6] := GVL_IO.bySafeOut6;
abySafeOut[7] := GVL_IO.bySafeOut7;

(* ============================================================================
   SIMULATION
   ============================================================================ *)

(* --- Call PROFIsafe simulator (Slot 1) --- *)
fbSafetySimulator(
    bEnable         := bSimulatorEnable,
    dwF_Source_Add  := dwF_Source_Add,
    dwF_Dest_Add    := dwF_Dest_Add,
    tF_WD_Time      := tF_WD_Time,
    abySafeOut      := abySafeOut,
    bCommOK         => bSafeCommOK
);

(* --- Call VASS simulator (Slot 2) with the program player --- *)
fbVassSimulator(
    bEnable         := bSimulatorEnable,
    wRobotID        := GVL_Program.ROBOT_INDEX,
    aVassOutputData := aVassOutputData,
    abySafeOut      := abySafeOut,
    rDt             := GVL_Program.R_TASK_S,
    bActive         => bSimActive,
    eCurrentMode    => eMode,
    eProgramState   => eProgState,
    bSafetyOK       => bSafetyHealthy
);
aVassInputData := fbVassSimulator.aVassInputData;
abySafeIn := fbVassSimulator.abySafeIn;
wActiveJob := fbVassSimulator.wActiveJob;
wCurrentStep := fbVassSimulator.wCurrentStep;
dwRequest := fbVassSimulator.dwRequest;
dwGrant := fbVassSimulator.dwGrant;
ePlayerState := fbVassSimulator.ePlayerState;

(* --- Joint angles from the player -> VASS Option area (bytes 16-27, big-endian) --- *)
fbJointEncoder(
    rA1_deg         := fbVassSimulator.rA1_deg,
    rA2_deg         := fbVassSimulator.rA2_deg,
    rA3_deg         := fbVassSimulator.rA3_deg,
    rA4_deg         := fbVassSimulator.rA4_deg,
    rA5_deg         := fbVassSimulator.rA5_deg,
    rA6_deg         := fbVassSimulator.rA6_deg
);
FOR _i := 0 TO 11 DO
    aVassInputData[16 + _i] := fbJointEncoder.abyOption[_i];
END_FOR

(* Monitor: decode back for quick verification in debug view *)
rMonitor_A1_deg := INT_TO_REAL(fbJointEncoder.iA1_count) * 0.02;
rMonitor_A2_deg := INT_TO_REAL(fbJointEncoder.iA2_count) * 0.02;
rMonitor_A3_deg := INT_TO_REAL(fbJointEncoder.iA3_count) * 0.02;
rMonitor_A4_deg := INT_TO_REAL(fbJointEncoder.iA4_count) * 0.02;
rMonitor_A5_deg := INT_TO_REAL(fbJointEncoder.iA5_count) * 0.02;
rMonitor_A6_deg := INT_TO_REAL(fbJointEncoder.iA6_count) * 0.02;

(* --- Debug: Error injection --- *)
(* Set bTest_InjectError := TRUE in online/debug view to simulate a robot error *)
IF bTest_InjectError THEN
    aVassInputData[0] := aVassInputData[0] OR BYTE#16#40;   (* Set bit 6 = Error *)
    aVassInputData[10] := WORD_TO_BYTE(wTest_ErrorCode AND WORD#16#FF);
    aVassInputData[11] := WORD_TO_BYTE(SHR(wTest_ErrorCode, 8));
END_IF

IF bTest_InjectSafetyFault THEN
    abySafeIn[2] := abySafeIn[2] OR BYTE#16#80;     (* Set bit 7 = Fault *)
    abySafeIn[0] := abySafeIn[0] AND BYTE#16#FE;    (* Clear bit 0 = Drives NOT OK *)
END_IF

(* ============================================================================
   OUTPUTS: write the robot status back to GVL_IO (whole array / scalars)
   ============================================================================ *)
GVL_IO.aVassInputData := aVassInputData;
GVL_IO.bySafeIn0 := abySafeIn[0];
GVL_IO.bySafeIn1 := abySafeIn[1];
GVL_IO.bySafeIn2 := abySafeIn[2];
GVL_IO.bySafeIn3 := abySafeIn[3];
GVL_IO.bySafeIn4 := abySafeIn[4];
GVL_IO.bySafeIn5 := abySafeIn[5];
GVL_IO.bySafeIn6 := abySafeIn[6];
GVL_IO.bySafeIn7 := abySafeIn[7];
